Fanuc KAREL source: kx00020.KL

PROGRAM KX00020
%NOLOCKGROUP
VAR
I:INTEGER;J:INTEGER;B:BOOLEAN
F : FILE
S : STRING[80]
P : XYZWPR
SA : ARRAY[4] OF STRING[12]
BEGIN
--
--
SA[1]='A'
S=SA[1]
END KX00020
